FUNCTION_BLOCK POSTGRE_DB_INSERT
  {SET_ATTRIBUTE(OpcUa, POINT.ENDPOINT)}
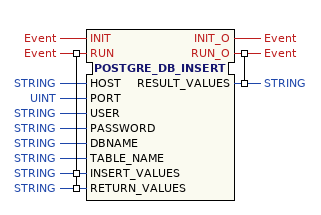
  EVENT_INPUT
    INIT;
    RUN WITH INSERT_VALUES, RETURN_VALUES;
  END_EVENT
  EVENT_OUTPUT
    INIT_O;
    RUN_O WITH RESULT_VALUES;
  END_EVENT
  VAR_INPUT
    HOST : STRING; {SET_ATTRIBUTE(OpcUa, Constant)}
    PORT : UINT; {SET_ATTRIBUTE(OpcUa, Constant)}
    USER : STRING; {SET_ATTRIBUTE(OpcUa, Constant)}
    PASSWORD : STRING; {SET_ATTRIBUTE(OpcUa, Constant)}
    DBNAME : STRING; {SET_ATTRIBUTE(OpcUa, Constant)}
    TABLE_NAME : STRING; {SET_ATTRIBUTE(OpcUa, Constant)}
    INSERT_VALUES : STRING; {SET_ATTRIBUTE(OpcUa, Variable.RUN)}
    RETURN_VALUES : STRING; {SET_ATTRIBUTE(OpcUa, Variable.RUN)}
  END_VAR
  VAR_OUTPUT
    RESULT_VALUES : STRING; {SET_ATTRIBUTE(OpcUa, Variable.RUN)}
  END_VAR
END_FUNCTION_BLOCK
